INTERFACE I_Parameters_MainControl

PROPERTY cylinderSensorTimeout : TIME
GET
END_GET
END_PROPERTY

PROPERTY isLoggerEnabled : BOOL
GET
END_GET
END_PROPERTY

PROPERTY numberOfRetries : INT
GET
END_GET
END_PROPERTY

END_INTERFACE

(* stored: Version 1.1.0.1, ProductVersion 3.1.4024.12
   Itf I_Parameters_MainControl: Id {ac418b51-b2c2-4e75-8392-0f9fe5c71974}
   Property cylinderSensorTimeout: Id {a539eef0-e668-4d30-bdf4-17d19fc50d5c}
   Get Get: Id {1d4b370b-eb35-4a73-91e4-c2a260391746}
   Property isLoggerEnabled: Id {24545445-dc74-42e9-b1c6-b3af94d10f62}
   Get Get: Id {8fc51ee9-5587-43fd-b626-46e233e7f3cb}
   Property numberOfRetries: Id {3250e2cb-c237-42a7-be55-e0c13f4e8e1e}
   Get Get: Id {240e4671-b07e-442b-95c3-d9f229abd2d8} *)
